FUNCTION_BLOCK FB_ExtTilt
(*

The function block used to generate move external trajectory.

Constructor: 		Patryk Panylo
Company:		E. Riexinger GmbH
Date:			01.04.2015
Version:			1.00

Date:			Revision:		Who:				Comment
dd.mm.yyyy		x.xx			Initials			comment

*)
VAR_INPUT
	(* Input variables / Eingang Variablen *)
	bEnable							:BOOL;						(* Function block enable *)
	bStart							:BOOL;						(* Execute start an external trajectory with rising edge *)
	bStop							:BOOL;						(* Execute stop an external trajectory with rising edge *)
	lrStartPosHorizontal				:LREAL;						(* Start position of horizontal axis [mm] *)
	lrStartPosVertical					:LREAL;						(* Start position of vertical axis [mm] *)
	lrOffsetPosHorizontal				:LREAL;						(* Offset position of horizontal axis [mm] *)
	lrOffsetPosVertical					:LREAL;						(* Offset position of vertical axis [mm] *)
	lrAngle							:LREAL;						(* Angle [°] *)
	unPosWindow					:UINT := 2;					(* Position window [mm] *)
	bTakeHorMovePara				:BOOL;						(* Take move parameters from 1- horizontal axis, 0 - vertical axis *)
END_VAR
VAR_OUTPUT
	(* Output variables / Ausgang Variablen *)
	lrNewPos						:LREAL;						(* New position [mm] *)
	lrNewVelo						:LREAL;						(* New velocity [mm/s] *)
	lrNewAcc						:LREAL;						(* New acceleration [mm/s^2] *)
	bEnabled  						:BOOL;						(* Calculate positon is enabled *)
	bDone							:BOOL;						(* Command done *)
	bBusy							:BOOL;						(* Command busy *)
	bError							:BOOL;						(* Command error  *)
	udnErrorNo						:UDINT;						(* Error number *)
	sErrorMsg						:STRING; 					(* Error message *)
END_VAR
VAR_IN_OUT
	AxisHorizontal					:AXIS_REF;					(* The AXIS_REF data type  is an interface between the PLC and the NC and contains axis information *)
	AxisVertical						:AXIS_REF;					(* The AXIS_REF data type  is an interface between the PLC and the NC and contains axis information *)
END_VAR
VAR
	(* Instances / Instanzen *)

	(* Enumerator  *)
	etCalcExtTiltState					:ET_CalcExtTiltState;								(* Current state *)

	(* General flags / Allgemeine Variablen *)
	lrExtStartPosHorizontal				:LREAL;
	lrExtStartPosVertical				:LREAL;
	lrExtAngle						:LREAL;
	lrCacheNewPos					:LREAL;						(* Cache new position [mm] *)
	bFirstTime						:BOOL;

END_VAR
VAR CONSTANT

END_VAR


IF NOT bEnable
THEN

	lrNewPos := SEL(bTakeHorMovePara, AxisVertical.NcToPlc.SetPos, AxisHorizontal.NcToPlc.SetPos);
	lrNewVelo := SEL(bTakeHorMovePara, AxisVertical.NcToPlc.SetVelo, AxisHorizontal.NcToPlc.SetVelo);
	lrNewAcc := SEL(bTakeHorMovePara, AxisVertical.NcToPlc.SetAcc, AxisHorizontal.NcToPlc.SetAcc);

	bDone := FALSE;					(* Command done *)
	bBusy := FALSE;					(* Command busy *)
	bError := FALSE;					(* Command error  *)
	udnErrorNo := 0;					(* Error number *)
	sErrorMsg := ''; 					(* Error message *)

	bEnabled := bStart;

	bFirstTime := FALSE;
	RETURN;
END_IF

IF NOT bFirstTime
THEN
	bEnabled := FALSE;

	etCalcExtTiltState := ET_CalcExtTiltState_eWaitExecute;

	bFirstTime := TRUE;
END_IF

CASE etCalcExtTiltState
OF
	ET_CalcExtTiltState_eWaitExecute:
		IF bStop
		THEN
			bEnabled := FALSE;

			bDone := FALSE;						(* Command done *)
			bBusy := TRUE;						(* Command busy *)
			bError := FALSE;						(* Command error  *)
			udnErrorNo := 0;						(* Error number *)
			sErrorMsg := ''; 						(* Error message *)

			etCalcExtTiltState := ET_CalcExtTiltState_eDone;

		ELSIF bStart
		THEN
			bDone := FALSE;						(* Command done *)
			bBusy := TRUE;						(* Command busy *)
			bError := FALSE;						(* Command error  *)
			udnErrorNo := 0;						(* Error number *)
			sErrorMsg := ''; 						(* Error message *)

			etCalcExtTiltState := ET_CalcExtTiltState_eCalcTiltPos;

		END_IF

	ET_CalcExtTiltState_eCalcTiltPos:
		bEnabled := TRUE;

		lrExtStartPosHorizontal := lrStartPosHorizontal;
		lrExtStartPosVertical := lrStartPosVertical;
		lrExtAngle := lrAngle;

		etCalcExtTiltState := ET_CalcExtTiltState_eDone;

	ET_CalcExtTiltState_eError:
		bBusy := FALSE;						(* Command busy *)
		bError := TRUE;						(* Command error  *)

		etCalcExtTiltState := ET_CalcExtTiltState_eNoExecute;

	ET_CalcExtTiltState_eDone:
		bDone := TRUE;						(* Command done *)
		bBusy := FALSE;						(* Command busy *)

		etCalcExtTiltState := ET_CalcExtTiltState_eNoExecute;

	ET_CalcExtTiltState_eNoExecute:
		IF NOT bStart
		     AND NOT bStop
		THEN
			(* Reset outputs *)
			bDone := FALSE;						(* Command done *)
			bBusy := FALSE;						(* Command busy *)
			bError := FALSE;						(* Command error  *)

			etCalcExtTiltState := ET_CalcExtTiltState_eWaitExecute;
		END_IF
END_CASE

(* The function is used to calculate a trajectory of vertical position. *)
IF bEnabled
THEN
	lrNewPos := F_CalcTiltPos(
		lrStartPosHorizontal := lrExtStartPosHorizontal,
		lrStartPosVertical := lrExtStartPosVertical,
		lrCurrentPosHorizontal := AxisHorizontal.NcToPlc.SetPos,
		lrCurrentPosVertical := AxisVertical.NcToPlc.SetPos,
		lrOffsetPosHorizontal := lrOffsetPosHorizontal,
		lrOffsetPosVertical := lrOffsetPosVertical,
		lrAngle :=lrExtAngle,
	);

	lrCacheNewPos := lrNewPos;
	lrNewVelo := AxisHorizontal.NcToPlc.SetVelo;
	lrNewAcc := AxisHorizontal.NcToPlc.SetAcc;

ELSE

	lrNewPos := SEL(bTakeHorMovePara, AxisVertical.NcToPlc.SetPos, AxisHorizontal.NcToPlc.SetPos);
	lrNewVelo := SEL(bTakeHorMovePara, AxisVertical.NcToPlc.SetVelo, AxisHorizontal.NcToPlc.SetVelo);
	lrNewAcc := SEL(bTakeHorMovePara, AxisVertical.NcToPlc.SetAcc, AxisHorizontal.NcToPlc.SetAcc);
	bError := FALSE;								(* Command error  *)
	udnErrorNo :=  0;								(* Error number *)
	sErrorMsg := ''; 								(* Error message *)
END_IF

END_FUNCTION_BLOCK

(* stored: Version 1.1.0.1, ProductVersion 3.1.4024.15
   POU FB_ExtTilt: Id {9df94794-92fa-449d-bcca-ef4314e6911f}, SpecialFunc None *)
